(* IEC 61131-3 sources: plc-vscode/tests/st/test-ready/trust-platform/examples/OSCAT/dairy_separator_adapter_state/non-oop/src, 3 files *)

(* ---- Main.st ---- *)
FUNCTION_BLOCK ClassicDairySeparator
VAR
    StateValue : INT;
    FeedValveOpenValue : BOOL;
    DischargeValveOpenValue : BOOL;
    CipValveOpenValue : BOOL;
    BowlRunningValue : BOOL;
    FaultCodeValue : DWORD;
END_VAR

METHOD PUBLIC Update : INT
VAR_INPUT
    StartCommand : BOOL;
    DischargeRequest : BOOL;
    CipMode : BOOL;
    UseSiemens : BOOL;
    StatusWord : WORD;
    SpeedFeedbackRpm : REAL;
    VibrationMmS : REAL;
    FaultRaw : WORD;
END_VAR
VAR
    RunningBit : BOOL;
    FaultBit : BOOL;
    AtSpeed : BOOL;
    VibrationHigh : BOOL;
END_VAR
IF UseSiemens THEN
    RunningBit := (WORD_TO_DWORD(StatusWord) AND DWORD#16#0400) <> DWORD#0;
    FaultCodeValue := DWORD#16#50000000 OR WORD_TO_DWORD(FaultRaw);
ELSE
    RunningBit := (WORD_TO_DWORD(StatusWord) AND DWORD#16#0004) <> DWORD#0;
    FaultCodeValue := DWORD#16#D0000000 OR WORD_TO_DWORD(FaultRaw);
END_IF;
FaultBit := (WORD_TO_DWORD(StatusWord) AND DWORD#16#0008) <> DWORD#0;
VibrationHigh := VibrationMmS > REAL#8.0;
AtSpeed := (SpeedFeedbackRpm >= REAL#6000.0) AND NOT FaultBit AND NOT VibrationHigh;

IF VibrationHigh THEN
    IF UseSiemens THEN
        FaultCodeValue := DWORD#16#500000F1;
    ELSE
        FaultCodeValue := DWORD#16#D00000F1;
    END_IF;
END_IF;

IF FaultBit OR VibrationHigh THEN
    StateValue := INT#90;
ELSIF StateValue = INT#0 THEN
    IF CipMode THEN
        StateValue := INT#40;
    ELSIF StartCommand THEN
        StateValue := INT#10;
    END_IF;
ELSIF StateValue = INT#10 THEN
    IF CipMode THEN
        StateValue := INT#40;
    ELSIF AtSpeed THEN
        StateValue := INT#20;
    END_IF;
ELSIF StateValue = INT#20 THEN
    IF CipMode THEN
        StateValue := INT#40;
    ELSIF DischargeRequest THEN
        StateValue := INT#30;
    ELSIF NOT AtSpeed THEN
        StateValue := INT#90;
    END_IF;
ELSIF StateValue = INT#30 THEN
    IF CipMode THEN
        StateValue := INT#40;
    ELSIF NOT DischargeRequest THEN
        StateValue := INT#20;
    END_IF;
ELSIF StateValue = INT#40 THEN
    IF NOT CipMode THEN
        StateValue := INT#0;
    END_IF;
END_IF;

FeedValveOpenValue := StateValue = INT#20;
DischargeValveOpenValue := StateValue = INT#30;
CipValveOpenValue := StateValue = INT#40;
BowlRunningValue := RunningBit OR (StateValue = INT#10) OR (StateValue = INT#20) OR (StateValue = INT#30);
Update := StateValue;
END_METHOD

PUBLIC PROPERTY FeedValveOpen : BOOL
GET
    FeedValveOpen := FeedValveOpenValue;
END_GET
END_PROPERTY

PUBLIC PROPERTY BowlRunning : BOOL
GET
    BowlRunning := BowlRunningValue;
END_GET
END_PROPERTY

PUBLIC PROPERTY FaultCode : DWORD
GET
    FaultCode := FaultCodeValue;
END_GET
END_PROPERTY
END_FUNCTION_BLOCK

PROGRAM Main
VAR
    Separator : ClassicDairySeparator;
    StartCommand : BOOL;
    DischargeRequest : BOOL;
    CipMode : BOOL;
    UseSiemensDrive : BOOL;
    StatusWordRaw : WORD;
    SpeedFeedbackRaw : INT;
    VibrationRaw : INT;
    FaultRaw : WORD;
    FeedValveOut : BOOL;
    DischargeValveOut : BOOL;
    CipValveOut : BOOL;
END_VAR
Separator.Update(StartCommand := StartCommand, DischargeRequest := DischargeRequest, CipMode := CipMode, UseSiemens := UseSiemensDrive, StatusWord := StatusWordRaw, SpeedFeedbackRpm := INT_TO_REAL(SpeedFeedbackRaw), VibrationMmS := INT_TO_REAL(VibrationRaw) / REAL#10.0, FaultRaw := FaultRaw);
FeedValveOut := Separator.FeedValveOpen;
DischargeValveOut := DischargeRequest;
CipValveOut := CipMode;
END_PROGRAM

(* ---- Configuration.st ---- *)
CONFIGURATION DairySeparatorAdapterStateClassicConfiguration
RESOURCE Cpu0 ON PLC
    TASK MainTask (INTERVAL := T#50ms, PRIORITY := 1);
    PROGRAM Separator WITH MainTask : Main;
END_RESOURCE
VAR_CONFIG
    Separator.StartCommand AT %IX0.0 : BOOL;
    Separator.DischargeRequest AT %IX0.1 : BOOL;
    Separator.CipMode AT %IX0.2 : BOOL;
    Separator.UseSiemensDrive AT %IX0.3 : BOOL;
    Separator.StatusWordRaw AT %IW0 : WORD;
    Separator.SpeedFeedbackRaw AT %IW2 : INT;
    Separator.VibrationRaw AT %IW4 : INT;
    Separator.FaultRaw AT %IW6 : WORD;
    Separator.FeedValveOut AT %QX0.0 : BOOL;
    Separator.DischargeValveOut AT %QX0.1 : BOOL;
    Separator.CipValveOut AT %QX0.2 : BOOL;
END_VAR
END_CONFIGURATION

(* ---- Tests.st ---- *)
TEST_PROGRAM ClassicSeparatorRunsProduction
VAR
    Separator : ClassicDairySeparator;
END_VAR

ASSERT_EQUAL(EXPECTED := INT#10, ACTUAL := Separator.Update(StartCommand := TRUE, DischargeRequest := FALSE, CipMode := FALSE, UseSiemens := FALSE, StatusWord := WORD#16#0004, SpeedFeedbackRpm := REAL#0.0, VibrationMmS := REAL#2.0, FaultRaw := WORD#16#0044));
ASSERT_EQUAL(EXPECTED := INT#20, ACTUAL := Separator.Update(StartCommand := TRUE, DischargeRequest := FALSE, CipMode := FALSE, UseSiemens := FALSE, StatusWord := WORD#16#0004, SpeedFeedbackRpm := REAL#6500.0, VibrationMmS := REAL#2.0, FaultRaw := WORD#16#0044));
ASSERT_TRUE(IN := Separator.FeedValveOpen);
END_TEST_PROGRAM

TEST_PROGRAM ClassicSeparatorTripsOnVibration
VAR
    Separator : ClassicDairySeparator;
END_VAR

ASSERT_EQUAL(EXPECTED := INT#90, ACTUAL := Separator.Update(StartCommand := TRUE, DischargeRequest := FALSE, CipMode := FALSE, UseSiemens := TRUE, StatusWord := WORD#16#0400, SpeedFeedbackRpm := REAL#6100.0, VibrationMmS := REAL#9.5, FaultRaw := WORD#16#0012));
ASSERT_EQUAL(EXPECTED := DWORD#16#500000F1, ACTUAL := Separator.FaultCode);
END_TEST_PROGRAM
